(* IEC 61131-3 sources: PLC-Static-Analysis/modules/plc-rules/src/test/resources/PLCA-L014, 2 files *)

(* ---- noncompliant.st ---- *)
FUNCTION_BLOCK FB_X
VAR_INPUT
    x : INT;
END_VAR
END_FUNCTION_BLOCK

PROGRAM P_L014
VAR
    n : INT;
    m : INT;
    r : REAL;
    b : BOOL;
    c : BOOL;
    q : BOOL;
    aData : ARRAY[1..3] OF INT;
    fbX : FB_X;
END_VAR
n := n; // PLCA-L014
aData[1] := aData[1]; // PLCA-L014
fbX.x := fbx.X; // PLCA-L014
END_PROGRAM

(* ---- compliant.st ---- *)
PROGRAM P_L014ok
VAR
    n : INT;
    m : INT;
    r : REAL;
    b : BOOL;
    c : BOOL;
    q : BOOL;
    aData : ARRAY[1..3] OF INT;
END_VAR
n := m;
n := n + 0;
aData[1] := aData[2];
END_PROGRAM
